// TIA Portal V21 export
// export: Created 2026-11-21T13:00:31.5652979Z, ExportSetting WithDefaults, DisplayName Totally Integrated Automation Portal, DisplayVersion V21, DisplayName STEP 7 Professional, DisplayVersion V21, DisplayName STEP 7 Safety, DisplayVersion V21, DisplayName Tech WebApplication, DisplayVersion V21, DisplayName WinCC Basic/Comfort/Advanced, DisplayVersion V21, DisplayName WinCC Unified, DisplayVersion V21
FUNCTION_BLOCK "Batch"   // FB20, GRAPH
TITLE = Batch sequence
VERSION : 0.1
// A batch sequence: fill and heat at once, mix, then drain or reject.
// stored: AcknowledgeErrorsRequired true, AutoNumber true, GraphVersion 6.0, InitialValuesAcquisition false, IsIECCheckEnabled false, LanguageInNetworks LAD, LockOperatingMode false, PermanentILProcessingInMANMode false, SetENOAutomatically false, SkipSteps false, UDAEnableTagReadback false, WithAlarmHandling true
   // inherited from GRAPH_BASE
   VAR
      OFF_SQ_BASE : Bool;
   END_VAR
   VAR_INPUT
      ACK_EF : Bool := false;   // Acknowledge all errors and faults
      start : Bool;
      full : Bool;
      hot : Bool;
      quality : Bool;
      door : Bool;
      overflow : Bool;
      acknowledge : Bool;
      level : Int;
   END_VAR
   VAR_OUTPUT
      valve : Bool;
      lamp : Bool;
      heater : Bool;
      mixer : Bool;
      drain : Bool;
      alarm : Bool;
      clamped : Int;
   END_VAR
BEGIN
// Sequence
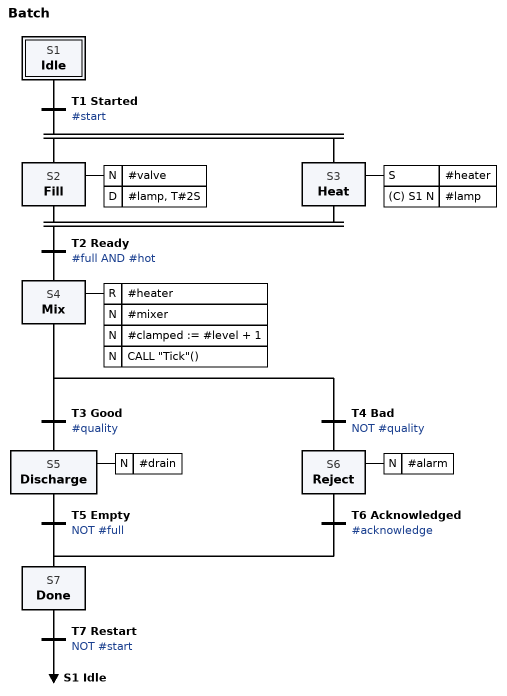
   // permanent pre-instructions
   NETWORK 1
      #lamp := #acknowledge;

   // sequencer 1
   INITIAL_STEP Idle:   // S1, max time T#10S, warning time T#7S
   END_STEP
   TRANSITION Started FROM Idle TO (Fill, Heat)   // T1
      := #start;
   END_TRANSITION
   STEP Fill:   // S2, max time T#10S, warning time T#7S
      supervision V := #overflow;
              N    #valve
              D    #lamp, T#2S
   END_STEP
   STEP Heat:   // S3, max time T#10S, warning time T#7S
      interlock C := #door;
              S    #heater
      (C) S1  N    #lamp
   END_STEP
   TRANSITION Ready FROM (Fill, Heat) TO Mix   // T2
      := #full AND #hot;
   END_TRANSITION
   STEP Mix:   // S4, max time T#10S, warning time T#7S
              R    #heater
              N    #mixer
              N    #clamped := #level + 1
              N    CALL "Tick"()
   END_STEP
   TRANSITION Good FROM Mix TO Discharge   // T3
      := #quality;
   END_TRANSITION
   TRANSITION Bad FROM Mix TO Reject   // T4
      := NOT #quality;
   END_TRANSITION
   STEP Discharge:   // S5, max time T#10S, warning time T#7S
              N    #drain
   END_STEP
   TRANSITION Empty FROM Discharge TO Done   // T5
      := NOT #full;
   END_TRANSITION
   STEP Reject:   // S6, max time T#10S, warning time T#7S
              N    #alarm
   END_STEP
   TRANSITION Acknowledged FROM Reject TO Done   // T6
      := #acknowledge;
   END_TRANSITION
   STEP Done:   // S7, max time T#10S, warning time T#7S
   END_STEP
   TRANSITION Restart FROM Done TO Idle   // T7, jump
      := NOT #start;
   END_TRANSITION

   // permanent post-instructions
   NETWORK 1
      #alarm := #overflow;
END_FUNCTION_BLOCK
